Fanuc KAREL source: KT00899.KL

PROGRAM KT00899
%NOLOCKGROUP
VAR
  P1: XYZWPR
  P2: XYZWPR
  OUT: BOOLEAN
BEGIN
  P1.X = 1.0
  P2.Y = 2.0
  P1.X = 1.0
  P2.Y = 2.0
  OUT = J_IN_RANGE(P1)
END KT00899
